FUNCTION_BLOCK GATE_CYCLE (* Migrated from IEC 61131-3 ST *)
  (* Standard: 61499-2 *)
  (* Version 1.0, 2026-11-06, st2fb *)
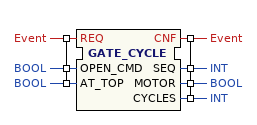
  EVENT_INPUT
    REQ WITH OPEN_CMD, AT_TOP;
  END_EVENT
  EVENT_OUTPUT
    CNF WITH SEQ, MOTOR, CYCLES;
  END_EVENT
  VAR_INPUT
    OPEN_CMD : BOOL;
    AT_TOP : BOOL;
  END_VAR
  VAR_OUTPUT
    SEQ : INT;
    MOTOR : BOOL;
    CYCLES : INT;
  END_VAR
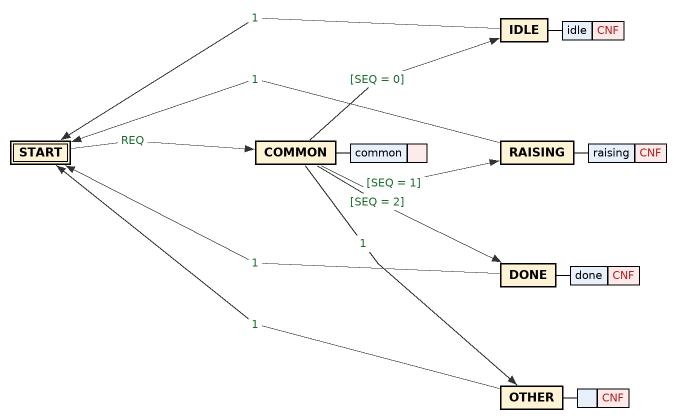
  EC_STATES
    START;
    COMMON : common;
    IDLE : idle -> CNF;
    RAISING : raising -> CNF;
    DONE : done -> CNF;
    OTHER : -> CNF;
  END_STATES
  EC_TRANSITIONS
    START TO COMMON := REQ;
    COMMON TO IDLE := [SEQ = 0];
    COMMON TO RAISING := [SEQ = 1];
    COMMON TO DONE := [SEQ = 2];
    COMMON TO OTHER := 1;
    IDLE TO START := 1;
    RAISING TO START := 1;
    DONE TO START := 1;
    OTHER TO START := 1;
  END_TRANSITIONS
  ALGORITHM common IN ST:
MOTOR := FALSE;
  END_ALGORITHM
  ALGORITHM idle IN ST:
IF OPEN_CMD THEN
  SEQ := 1;
END_IF;
  END_ALGORITHM
  ALGORITHM raising IN ST:
MOTOR := TRUE;
IF AT_TOP THEN
  SEQ := 2;
END_IF;
  END_ALGORITHM
  ALGORITHM done IN ST:
CYCLES := CYCLES + 1;
SEQ := 0;
  END_ALGORITHM
END_FUNCTION_BLOCK
